Fanuc KAREL source: KO00134.KL

PROGRAM KO00134
%NOLOCKGROUP
VAR
  R: REAL
  CFG: CONFIG
  OUT: XYZWPR
  N: REAL
BEGIN
  N = 1
  R = 2.0
  CFG.CFG_FLIP = TRUE
  OUT = POS(R, N, R, R, R, R, CFG)
END KO00134
